FUNCTION_BLOCK FB_CoverStoppingState EXTENDS FB_CoverState
VAR_INPUT
END_VAR
VAR_OUTPUT
END_VAR
VAR
END_VAR

METHOD RunState : BOOL
// Stop Motor 1
pCover^._Motor1RelaisA := FALSE;
pCover^._Motor1RelaisB := FALSE;
// Stop Motor 2
pCover^._Motor2RelaisA := FALSE;
pCover^._Motor2RelaisB := FALSE;
THIS^.SuccessfulFinished();
END_METHOD

METHOD SuccessfulFinished : BOOL
pCover^._CoverState := E_MirrorCoverState.stopped;
pCover^.SetState(pCover^.fbCoverIdleState);
END_METHOD

END_FUNCTION_BLOCK

(* stored: Version 1.1.0.1, ProductVersion 3.1.4024.15
   POU FB_CoverStoppingState: Id {f48b8b07-47c1-4266-826f-5feb1ff6fbca}, SpecialFunc None
   Method RunState: Id {7fdd173a-4c60-45f6-b8c9-8d404fcf0de6}
   Method SuccessfulFinished: Id {16696f42-d127-4d1e-b50e-ff1289983df1} *)
